// TIA Portal V19 export
DATA_BLOCK "RAMP_DB"   // DB11
// stored: InstanceOfName RAMP, InstanceOfType FB
"RAMP"
   // VAR_INPUT
   //    RAMP_START : Bool;
   //    JACKET_TT02 : Real;
   //    MASS_TT03 : Real;
   //    PRODUCT_TT : Real;
   //    RESET : Bool;
   //    SP : Real;
   //    PV : Real;
   //    "TIME" : Int;
   //    MAIN_START : Bool;
   //    MAIN_TIME : Int;
   //    MAIN_RESET : Bool;
   //    JACKET : Bool;
   //    MASS : Bool;
   //    PRODUCT : Bool;
   //    "A/M" : Bool;
   //    TIMER_RESET : Bool;
   //    COOL_RUNNING : Bool;
   //    HEAT_RUUNNING : Bool;
   //    SEMI : Bool;
   // END_VAR
   // VAR_OUTPUT
   //    RAMP_SP : Real;
   //    RAMP_RATE : Real;
   //    MAIN_COM : Bool;
   //    MAIN_PV : Real;
   //    RAMP_MIN : Int;
   // END_VAR
   // VAR_IN_OUT
   //    RAMP_INPUT : Real;
   //    TIME_1 : Int;
   //    ramp_substitute : Real;
   // END_VAR
   // VAR
   //    RampFunction_Instance { S7_SetPoint := 'True'} : RampFunction;
   //    TIMER_SECONDS_Instance { S7_SetPoint := 'True'} : "TIMER_SECONDS";
   //    START_MAIN_TIMER { S7_SetPoint := 'True'} : Bool;
   //    RAMP_TEMP_OUT : Real;
   //    TIMER_SECONDS_Instance_1 { S7_SetPoint := 'True'} : "TIMER_SECONDS";
   //    RAMP_CV_CTL { S7_SetPoint := 'True'} : PID_Compact;
   //    PID_Compact_1 { S7_SetPoint := 'True'} : PID_Compact;
   //    NORM_MIN : Int;
   //    NORM_MAX : Int;
   //    SCALE_MIN : Real;
   //    SCALE_MAX : Real;
   //    MAN_INPUT : Int;
   //    NORM_OUT : Real;
   //    SCVOUT : Int;
   //    MANOUT : Int;
   //    AO : Int;
   //    TIMER_SECONDS_Instance_2 { S7_SetPoint := 'True'} : "TIMER_SECONDS";
   //    P_TRIG6 { S7_SetPoint := 'True'} : Bool;
   //    P_TRIG7 : Bool;
   //    SEC : Int;
   //    IEC_Timer_0_Instance { S7_SetPoint := 'True'} : TOF_TIME;
   //    IEC_Timer_0_Instance_1 { S7_SetPoint := 'True'} : TP_TIME;
   // END_VAR
BEGIN
END_DATA_BLOCK
